FUNCTION_BLOCK CASE_SEQUENCER (* Migrated from IEC 61131-3 ST *)
  (* Standard: 61499-2 *)
  (* Version 1.0, 2026-11-06, st2fb *)
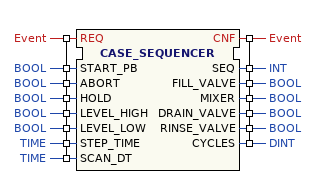
  EVENT_INPUT
    REQ WITH START_PB, ABORT, HOLD, LEVEL_HIGH, LEVEL_LOW, STEP_TIME, SCAN_DT;
  END_EVENT
  EVENT_OUTPUT
    CNF WITH SEQ, FILL_VALVE, MIXER, DRAIN_VALVE, RINSE_VALVE, CYCLES;
  END_EVENT
  VAR_INPUT
    START_PB : BOOL;
    ABORT : BOOL;
    HOLD : BOOL;
    LEVEL_HIGH : BOOL;
    LEVEL_LOW : BOOL;
    STEP_TIME : TIME;
    SCAN_DT : TIME;
  END_VAR
  VAR_OUTPUT
    SEQ : INT;
    FILL_VALVE : BOOL;
    MIXER : BOOL;
    DRAIN_VALVE : BOOL;
    RINSE_VALVE : BOOL;
    CYCLES : DINT;
  END_VAR
  VAR
    TIMING : BOOL;
    STEP_TIMER_IN : BOOL;
    STEP_TIMER_PT : TIME := T#0s;
    STEP_TIMER_Q : BOOL;
    STEP_TIMER_ET : TIME := T#0s;
    STEP_TIMER_STATE : INT := 0;
    STEP_TIMER_PREV_IN : BOOL;
    STEP_TIMER_START_TIME : TIME := T#0s;
    ST2FB_NOW : TIME := T#0s;
  END_VAR
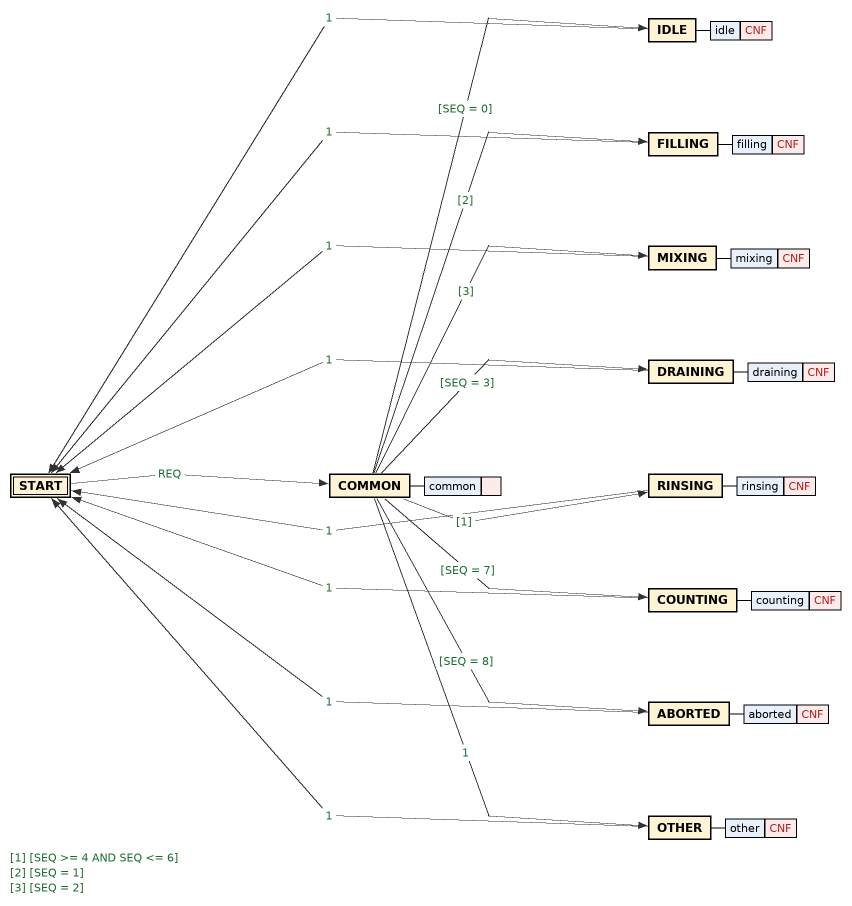
  EC_STATES
    START;
    COMMON : common;
    IDLE : idle -> CNF;
    FILLING : filling -> CNF;
    MIXING : mixing -> CNF;
    DRAINING : draining -> CNF;
    RINSING : rinsing -> CNF;
    COUNTING : counting -> CNF;
    ABORTED : aborted -> CNF;
    OTHER : other -> CNF;
  END_STATES
  EC_TRANSITIONS
    START TO COMMON := REQ;
    COMMON TO IDLE := [SEQ = 0];
    COMMON TO FILLING := [SEQ = 1];
    COMMON TO MIXING := [SEQ = 2];
    COMMON TO DRAINING := [SEQ = 3];
    COMMON TO RINSING := [SEQ >= 4 AND SEQ <= 6];
    COMMON TO COUNTING := [SEQ = 7];
    COMMON TO ABORTED := [SEQ = 8];
    COMMON TO OTHER := 1;
    IDLE TO START := 1;
    FILLING TO START := 1;
    MIXING TO START := 1;
    DRAINING TO START := 1;
    RINSING TO START := 1;
    COUNTING TO START := 1;
    ABORTED TO START := 1;
    OTHER TO START := 1;
  END_TRANSITIONS
  ALGORITHM common IN ST:
ST2FB_NOW := ST2FB_NOW + SCAN_DT;
IF NOT HOLD THEN
  STEP_TIMER_IN := TIMING;
  STEP_TIMER_PT := STEP_TIME;
  IF (STEP_TIMER_STATE = 0) AND NOT STEP_TIMER_PREV_IN AND STEP_TIMER_IN THEN
    STEP_TIMER_STATE := 1;
    STEP_TIMER_Q := FALSE;
    STEP_TIMER_START_TIME := ST2FB_NOW;
  ELSE
    IF NOT STEP_TIMER_IN THEN
      STEP_TIMER_ET := T#0s;
      STEP_TIMER_Q := FALSE;
      STEP_TIMER_STATE := 0;
    ELSIF STEP_TIMER_STATE = 1 THEN
      IF STEP_TIMER_START_TIME + STEP_TIMER_PT <= ST2FB_NOW THEN
        STEP_TIMER_STATE := 2;
        STEP_TIMER_Q := TRUE;
        STEP_TIMER_ET := STEP_TIMER_PT;
      ELSE
        STEP_TIMER_ET := ST2FB_NOW - STEP_TIMER_START_TIME;
      END_IF;
    END_IF;
  END_IF;
  STEP_TIMER_PREV_IN := STEP_TIMER_IN;
END_IF;
FILL_VALVE := FALSE;
MIXER := FALSE;
DRAIN_VALVE := FALSE;
RINSE_VALVE := FALSE;
IF ABORT THEN
  SEQ := 8;
END_IF;
  END_ALGORITHM
  ALGORITHM idle IN ST:
TIMING := FALSE;
IF START_PB THEN
  SEQ := 1;
END_IF;
  END_ALGORITHM
  ALGORITHM filling IN ST:
FILL_VALVE := TRUE;
IF LEVEL_HIGH THEN
  SEQ := 2;
  TIMING := TRUE;
END_IF;
  END_ALGORITHM
  ALGORITHM mixing IN ST:
MIXER := TRUE;
IF STEP_TIMER_Q THEN
  SEQ := 3;
  TIMING := FALSE;
END_IF;
  END_ALGORITHM
  ALGORITHM draining IN ST:
DRAIN_VALVE := TRUE;
IF LEVEL_LOW THEN
  SEQ := 4;
END_IF;
  END_ALGORITHM
  ALGORITHM rinsing IN ST:
RINSE_VALVE := TRUE;
IF STEP_TIMER_Q THEN
  SEQ := SEQ + 1;
  TIMING := FALSE;
ELSE
  TIMING := TRUE;
END_IF;
  END_ALGORITHM
  ALGORITHM counting IN ST:
CYCLES := CYCLES + 1;
SEQ := 0;
  END_ALGORITHM
  ALGORITHM aborted IN ST:
TIMING := FALSE;
DRAIN_VALVE := TRUE;
IF LEVEL_LOW AND NOT ABORT THEN
  SEQ := 0;
END_IF;
  END_ALGORITHM
  ALGORITHM other IN ST:
SEQ := 0;
  END_ALGORITHM
END_FUNCTION_BLOCK
